TYPE BodyMotion :
STRUCT
	distanceInM : LREAL;
	headingChangeInRad : LREAL;
END_STRUCT
END_TYPE

(* stored: Version 1.1.0.1, ProductVersion 3.1.4026.12
   DUT BodyMotion: Id {6f721b41-2435-54e2-9063-dbf309e6ec40} *)
